(* PLC project GeneratedProgram, SafePLC-Gen SafePLC-Gen Multimodal 1.0 *)
(* stored: creationDateTime 2026-04-25T11:49:46.044727Z *)

PROGRAM GeneratedProgram
  VAR
    FirstScan : BOOL;
    TICSA_4750_03_Scaled : REAL;
    PICSA_4712_02_Scaled : REAL;
    PI_4712_01_Scaled : REAL;
    TICSA_4750_03_SP : REAL;
    TICSA_4750_03_HH_SP : REAL;
    TICSA_4750_03_H_SP : REAL;
    TICSA_4750_03_L_SP : REAL;
    TICSA_4750_03_LL_SP : REAL;
    TICSA_4750_03_Deadband : REAL;
    TICSA_4750_03_H : BOOL;
    TICSA_4750_03_L : BOOL;
    TICSA_4750_03_HH_Latch : SR;
    TICSA_4750_03_LL_Latch : SR;
    TICSA_4750_03_HH_Ack : BOOL;
    TICSA_4750_03_LL_Ack : BOOL;
    PICSA_4712_02_SP : REAL;
    PICSA_4712_02_HH_SP : REAL;
    PICSA_4712_02_H_SP : REAL;
    PICSA_4712_02_L_SP : REAL;
    PICSA_4712_02_LL_SP : REAL;
    PICSA_4712_02_Deadband : REAL;
    PICSA_4712_02_H : BOOL;
    PICSA_4712_02_L : BOOL;
    PICSA_4712_02_HH_Latch : SR;
    PICSA_4712_02_LL_Latch : SR;
    PICSA_4712_02_HH_Ack : BOOL;
    PICSA_4712_02_LL_Ack : BOOL;
    PI_4712_01_HH_SP : REAL;
    PI_4712_01_H_SP : REAL;
    PI_4712_01_L_SP : REAL;
    PI_4712_01_LL_SP : REAL;
    PI_4712_01_Deadband : REAL;
    PI_4712_01_H : BOOL;
    PI_4712_01_L : BOOL;
    PI_4712_01_HH_Latch : SR;
    PI_4712_01_LL_Latch : SR;
    PI_4712_01_HH_Ack : BOOL;
    PI_4712_01_LL_Ack : BOOL;
    LOOP_4750_03_TRIP : BOOL;
    LOOP_4712_02_TRIP : BOOL;
    LOOP_104_01_TRIP : BOOL;
    TICSA_4750_03_HH : BOOL;
    TICSA_4750_03_LL : BOOL;
    PICSA_4712_02_HH : BOOL;
    PICSA_4712_02_LL : BOOL;
    SV_104_01_HH : BOOL;
    SV_104_01_LL : BOOL;
    SAFE_STATE : BOOL;
    TIC_Error : REAL;
    TIC_Integral : REAL;
    TIC_Kp : REAL;
    TIC_Ki : REAL;
    TIC_Output : REAL;
    PIC_Error : REAL;
    PIC_Integral : REAL;
    PIC_Kp : REAL;
    PIC_Ki : REAL;
    PIC_Output : REAL;
    SV_104_01_Out : BOOL;
    HV_MNb_47123_ISO_Out : BOOL;
    CHK_73KH12_50_P4712_Out : BOOL;
    CHK_MNc_47124_P4712_Out : BOOL;
    STR_75SA21_80_Out : BOOL;
    BV_75HB13_73HG12_Out : BOOL;
    BV_Q_80_N6_Out : BOOL;
    HV_QSa_47140_Out : BOOL;
    HV_QSb_47141_Out : BOOL;
    SB_Q_80_N6_Out : BOOL;
    System_Alarm : BOOL;
  END_VAR

            IF FirstScan THEN
    LOOP_4750_03_TRIP := TRUE;
    LOOP_4712_02_TRIP := TRUE;
    LOOP_104_01_TRIP  := TRUE;
    SAFE_STATE        := TRUE;
    TV_4750_03_Out    := 32767;
    PV_4712_02_Out    := 6554;
    XV_4750_01        := FALSE;
    SV_104_01_Out              := FALSE;
    HV_MNb_47123_ISO_Out       := FALSE;
    CHK_73KH12_50_P4712_Out    := FALSE;
    CHK_MNc_47124_P4712_Out    := FALSE;
    STR_75SA21_80_Out          := FALSE;
    BV_75HB13_73HG12_Out       := FALSE;
    BV_Q_80_N6_Out             := FALSE;
    HV_QSa_47140_Out           := FALSE;
    HV_QSb_47141_Out           := FALSE;
    SB_Q_80_N6_Out             := FALSE;
    FirstScan         := FALSE;
    RETURN;
END_IF;

TICSA_4750_03_Scaled := ((INT_TO_REAL(TICSA_4750_03_Raw) - 6554.0) / (32767.0 - 6554.0)) * 150.0;
PICSA_4712_02_Scaled := ((INT_TO_REAL(PICSA_4712_02_Raw) - 6554.0) / (32767.0 - 6554.0)) * 10.0;
PI_4712_01_Scaled    := ((INT_TO_REAL(PI_4712_01_Raw)    - 6554.0) / (32767.0 - 6554.0)) * 10.0;

TICSA_4750_03_HH := TICSA_4750_03_Scaled > TICSA_4750_03_HH_SP;
TICSA_4750_03_LL := TICSA_4750_03_Scaled < TICSA_4750_03_LL_SP;
PICSA_4712_02_HH := PICSA_4712_02_Scaled > PICSA_4712_02_HH_SP;
PICSA_4712_02_LL := PICSA_4712_02_Scaled < PICSA_4712_02_LL_SP;
SV_104_01_HH     := HS_4750_01;
SV_104_01_LL     := FALSE;

IF TICSA_4750_03_HH OR TICSA_4750_03_LL THEN
    LOOP_4750_03_TRIP := TRUE;
ELSIF LOOP_4750_03_TRIP AND MANUAL_RESET
      AND NOT TICSA_4750_03_HH AND NOT TICSA_4750_03_LL THEN
    LOOP_4750_03_TRIP := FALSE;
END_IF;

IF PICSA_4712_02_HH OR PICSA_4712_02_LL THEN
    LOOP_4712_02_TRIP := TRUE;
ELSIF LOOP_4712_02_TRIP AND MANUAL_RESET
      AND NOT PICSA_4712_02_HH AND NOT PICSA_4712_02_LL THEN
    LOOP_4712_02_TRIP := FALSE;
END_IF;

IF SV_104_01_HH OR SV_104_01_LL THEN
    LOOP_104_01_TRIP := TRUE;
ELSIF LOOP_104_01_TRIP AND MANUAL_RESET
      AND NOT SV_104_01_HH AND NOT SV_104_01_LL THEN
    LOOP_104_01_TRIP := FALSE;
END_IF;

SAFE_STATE := ESTOP
              OR LOOP_4750_03_TRIP
              OR LOOP_4712_02_TRIP
              OR LOOP_104_01_TRIP;

IF NOT SAFE_STATE THEN
    TIC_Error    := TICSA_4750_03_SP - TICSA_4750_03_Scaled;
    TIC_Integral := TIC_Integral + (TIC_Ki * TIC_Error);
    IF TIC_Integral > 100.0 THEN
        TIC_Integral := 100.0;
    ELSIF TIC_Integral < 0.0 THEN
        TIC_Integral := 0.0;
    END_IF;
    TIC_Output := (TIC_Kp * TIC_Error) + TIC_Integral;
    IF TIC_Output > 100.0 THEN
        TIC_Output := 100.0;
    ELSIF TIC_Output < 0.0 THEN
        TIC_Output := 0.0;
    END_IF;
    TV_4750_03_Out := REAL_TO_INT(6554.0 + (TIC_Output / 100.0) * (32767.0 - 6554.0));
ELSE
    TV_4750_03_Out := 32767;
END_IF;

IF NOT SAFE_STATE THEN
    PIC_Error    := PICSA_4712_02_SP - PICSA_4712_02_Scaled;
    PIC_Integral := PIC_Integral + (PIC_Ki * PIC_Error);
    IF PIC_Integral > 100.0 THEN
        PIC_Integral := 100.0;
    ELSIF PIC_Integral < 0.0 THEN
        PIC_Integral := 0.0;
    END_IF;
    PIC_Output := (PIC_Kp * PIC_Error) + PIC_Integral;
    IF PIC_Output > 100.0 THEN
        PIC_Output := 100.0;
    ELSIF PIC_Output < 0.0 THEN
        PIC_Output := 0.0;
    END_IF;
    PV_4712_02_Out := REAL_TO_INT(6554.0 + (PIC_Output / 100.0) * (32767.0 - 6554.0));
ELSE
    PV_4712_02_Out := 6554;
END_IF;

IF NOT SAFE_STATE AND HS_4750_01 THEN
    XV_4750_01 := TRUE;
ELSE
    XV_4750_01 := FALSE;
END_IF;

IF NOT SAFE_STATE THEN
    SV_104_01_Out            := TRUE;
    HV_MNb_47123_ISO_Out     := TRUE;
    CHK_73KH12_50_P4712_Out  := TRUE;
    CHK_MNc_47124_P4712_Out  := TRUE;
    STR_75SA21_80_Out        := TRUE;
    BV_75HB13_73HG12_Out     := TRUE;
    BV_Q_80_N6_Out           := TRUE;
    HV_QSa_47140_Out         := TRUE;
    HV_QSb_47141_Out         := TRUE;
    SB_Q_80_N6_Out           := TRUE;
ELSE
    SV_104_01_Out            := FALSE;
    HV_MNb_47123_ISO_Out     := FALSE;
    CHK_73KH12_50_P4712_Out  := FALSE;
    CHK_MNc_47124_P4712_Out  := FALSE;
    STR_75SA21_80_Out        := FALSE;
    BV_75HB13_73HG12_Out     := FALSE;
    BV_Q_80_N6_Out           := FALSE;
    HV_QSa_47140_Out         := FALSE;
    HV_QSb_47141_Out         := FALSE;
    SB_Q_80_N6_Out           := FALSE;
END_IF;

(* Four-level alarms — TICSA-4750.03 *)
IF TICSA_4750_03_Scaled > TICSA_4750_03_HH_SP THEN
    TICSA_4750_03_HH_Latch.S1 := TRUE;
ELSIF TICSA_4750_03_Scaled <= (TICSA_4750_03_HH_SP - TICSA_4750_03_Deadband) THEN
    TICSA_4750_03_HH_Latch.S1 := FALSE;
END_IF;
TICSA_4750_03_HH_Latch.R := TICSA_4750_03_HH_Ack AND NOT TICSA_4750_03_HH;
TICSA_4750_03_HH_Latch(S1 := TICSA_4750_03_HH_Latch.S1, R := TICSA_4750_03_HH_Latch.R);

IF TICSA_4750_03_Scaled > TICSA_4750_03_H_SP THEN
    TICSA_4750_03_H := TRUE;
ELSIF TICSA_4750_03_Scaled <= (TICSA_4750_03_H_SP - TICSA_4750_03_Deadband) THEN
    TICSA_4750_03_H := FALSE;
END_IF;

IF TICSA_4750_03_Scaled < TICSA_4750_03_L_SP THEN
    TICSA_4750_03_L := TRUE;
ELSIF TICSA_4750_03_Scaled >= (TICSA_4750_03_L_SP + TICSA_4750_03_Deadband) THEN
    TICSA_4750_03_L := FALSE;
END_IF;

IF TICSA_4750_03_Scaled < TICSA_4750_03_LL_SP THEN
    TICSA_4750_03_LL_Latch.S1 := TRUE;
ELSIF TICSA_4750_03_Scaled >= (TICSA_4750_03_LL_SP + TICSA_4750_03_Deadband) THEN
    TICSA_4750_03_LL_Latch.S1 := FALSE;
END_IF;
TICSA_4750_03_LL_Latch.R := TICSA_4750_03_LL_Ack AND NOT TICSA_4750_03_LL;
TICSA_4750_03_LL_Latch(S1 := TICSA_4750_03_LL_Latch.S1, R := TICSA_4750_03_LL_Latch.R);

(* Four-level alarms — PICSA-4712.02 *)
IF PICSA_4712_02_Scaled > PICSA_4712_02_HH_SP THEN
    PICSA_4712_02_HH_Latch.S1 := TRUE;
ELSIF PICSA_4712_02_Scaled <= (PICSA_4712_02_HH_SP - PICSA_4712_02_Deadband) THEN
    PICSA_4712_02_HH_Latch.S1 := FALSE;
END_IF;
PICSA_4712_02_HH_Latch.R := PICSA_4712_02_HH_Ack AND NOT PICSA_4712_02_HH;
PICSA_4712_02_HH_Latch(S1 := PICSA_4712_02_HH_Latch.S1, R := PICSA_4712_02_HH_Latch.R);

IF PICSA_4712_02_Scaled > PICSA_4712_02_H_SP THEN
    PICSA_4712_02_H := TRUE;
ELSIF PICSA_4712_02_Scaled <= (PICSA_4712_02_H_SP - PICSA_4712_02_Deadband) THEN
    PICSA_4712_02_H := FALSE;
END_IF;

IF PICSA_4712_02_Scaled < PICSA_4712_02_L_SP THEN
    PICSA_4712_02_L := TRUE;
ELSIF PICSA_4712_02_Scaled >= (PICSA_4712_02_L_SP + PICSA_4712_02_Deadband) THEN
    PICSA_4712_02_L := FALSE;
END_IF;

IF PICSA_4712_02_Scaled < PICSA_4712_02_LL_SP THEN
    PICSA_4712_02_LL_Latch.S1 := TRUE;
ELSIF PICSA_4712_02_Scaled >= (PICSA_4712_02_LL_SP + PICSA_4712_02_Deadband) THEN
    PICSA_4712_02_LL_Latch.S1 := FALSE;
END_IF;
PICSA_4712_02_LL_Latch.R := PICSA_4712_02_LL_Ack AND NOT PICSA_4712_02_LL;
PICSA_4712_02_LL_Latch(S1 := PICSA_4712_02_LL_Latch.S1, R := PICSA_4712_02_LL_Latch.R);

(* Four-level alarms — PI-4712.01 *)
IF PI_4712_01_Scaled > PI_4712_01_HH_SP THEN
    PI_4712_01_HH_Latch.S1 := TRUE;
ELSIF PI_4712_01_Scaled <= (PI_4712_01_HH_SP - PI_4712_01_Deadband) THEN
    PI_4712_01_HH_Latch.S1 := FALSE;
END_IF;
PI_4712_01_HH_Latch.R := PI_4712_01_HH_Ack AND NOT (PI_4712_01_Scaled > PI_4712_01_HH_SP);
PI_4712_01_HH_Latch(S1 := PI_4712_01_HH_Latch.S1, R := PI_4712_01_HH_Latch.R);

IF PI_4712_01_Scaled > PI_4712_01_H_SP THEN
    PI_4712_01_H := TRUE;
ELSIF PI_4712_01_Scaled <= (PI_4712_01_H_SP - PI_4712_01_Deadband) THEN
    PI_4712_01_H := FALSE;
END_IF;

IF PI_4712_01_Scaled < PI_4712_01_L_SP THEN
    PI_4712_01_L := TRUE;
ELSIF PI_4712_01_Scaled >= (PI_4712_01_L_SP + PI_4712_01_Deadband) THEN
    PI_4712_01_L := FALSE;
END_IF;

IF PI_4712_01_Scaled < PI_4712_01_LL_SP THEN
    PI_4712_01_LL_Latch.S1 := TRUE;
ELSIF PI_4712_01_Scaled >= (PI_4712_01_LL_SP + PI_4712_01_Deadband) THEN
    PI_4712_01_LL_Latch.S1 := FALSE;
END_IF;
PI_4712_01_LL_Latch.R := PI_4712_01_LL_Ack AND NOT (PI_4712_01_Scaled < PI_4712_01_LL_SP);
PI_4712_01_LL_Latch(S1 := PI_4712_01_LL_Latch.S1, R := PI_4712_01_LL_Latch.R);

System_Alarm :=
    TICSA_4750_03_HH_Latch.Q1 OR TICSA_4750_03_LL_Latch.Q1 OR
    TICSA_4750_03_H            OR TICSA_4750_03_L            OR
    PICSA_4712_02_HH_Latch.Q1 OR PICSA_4712_02_LL_Latch.Q1 OR
    PICSA_4712_02_H            OR PICSA_4712_02_L            OR
    PI_4712_01_HH_Latch.Q1    OR PI_4712_01_LL_Latch.Q1    OR
    PI_4712_01_H               OR PI_4712_01_L               OR
    LOOP_4750_03_TRIP          OR LOOP_4712_02_TRIP          OR
    LOOP_104_01_TRIP           OR SAFE_STATE;
          
END_PROGRAM

CONFIGURATION Config0
  RESOURCE Res0 ON PLC
    TASK MainTask(INTERVAL := T#20ms, PRIORITY := 0);
    PROGRAM Main : GeneratedProgram;
  END_RESOURCE
END_CONFIGURATION
